FUNCTION_BLOCK AckHelper (* Basic Function Block Type *)
  (* Standard: 61499-2 *)
  (* Version 0.0, 10/22/2026, macie, Schneider Electric, Template *)
  PACKAGE Main;
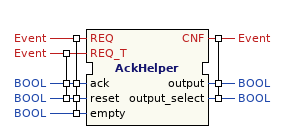
  EVENT_INPUT
    REQ WITH ack, reset, empty; (* Normal Execution Request *)
    REQ_T WITH ack, reset;
  END_EVENT
  EVENT_OUTPUT
    CNF WITH output, output_select; (* Execution Confirmation *)
  END_EVENT
  VAR_INPUT
    ack : BOOL; (* Input event qualifier *)
    reset : BOOL;
    empty : BOOL;
  END_VAR
  VAR_OUTPUT
    output : BOOL; (* Output event qualifier *)
    output_select : BOOL;
  END_VAR
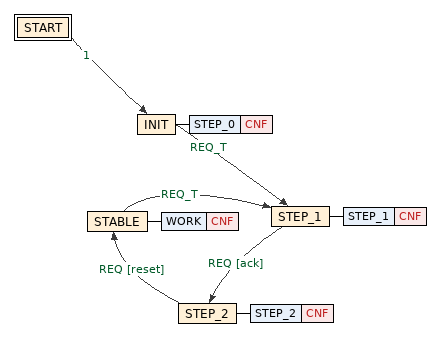
  EC_STATES
    START; (* Initial State *)
    INIT : STEP_0 -> CNF;
    STEP_1 : STEP_1 -> CNF;
    STEP_2 : STEP_2 -> CNF;
    STABLE : WORK -> CNF;
  END_STATES
  EC_TRANSITIONS
    START TO INIT := 1;
    INIT TO STEP_1 := REQ_T;
    STEP_1 TO STEP_2 := REQ [ack];
    STEP_2 TO STABLE := REQ [reset];
    STABLE TO STEP_1 := REQ_T;
  END_TRANSITIONS
  ALGORITHM STEP_0 IN ST: (* Normally executed algorithm *)
;
output := TRUE;
output_select := FALSE;
  END_ALGORITHM
  ALGORITHM STEP_1 IN ST:
;
output_select := TRUE;
  END_ALGORITHM
  ALGORITHM STEP_2 IN ST:
;
output := FALSE;
output_select := FALSE;
  END_ALGORITHM
  ALGORITHM WORK IN ST:
;
output := empty;
  END_ALGORITHM
END_FUNCTION_BLOCK
